FUNCTION FC 1 : VOID
BEGIN
NETWORK
      L MW 70000
END_FUNCTION
